// CFC twin of T_SafeOr_Tests: the same tests drawn as CFC diagrams, the way a TwinSAFE project is authored.
    FUNCTION_BLOCK T_SafeOr_Tests_CFC EXTENDS T_SafeCfcTestSuite
    VAR
    // Test_AnyConnectedInputTrueGivesRun
    group_1 : T_SafeGroup;
    fb_1 : T_SafeOr(group := group_1);
    // Test_AllFalseGivesSafe
    group_2 : T_SafeGroup;
    fb_2 : T_SafeOr(group := group_2);
END_VAR

Test_AnyConnectedInputTrueGivesRun();
Test_AllFalseGivesSafe();

METHOD PRIVATE Test_AnyConnectedInputTrueGivesRun
// note: this text did not pass the execution check against the stored diagram
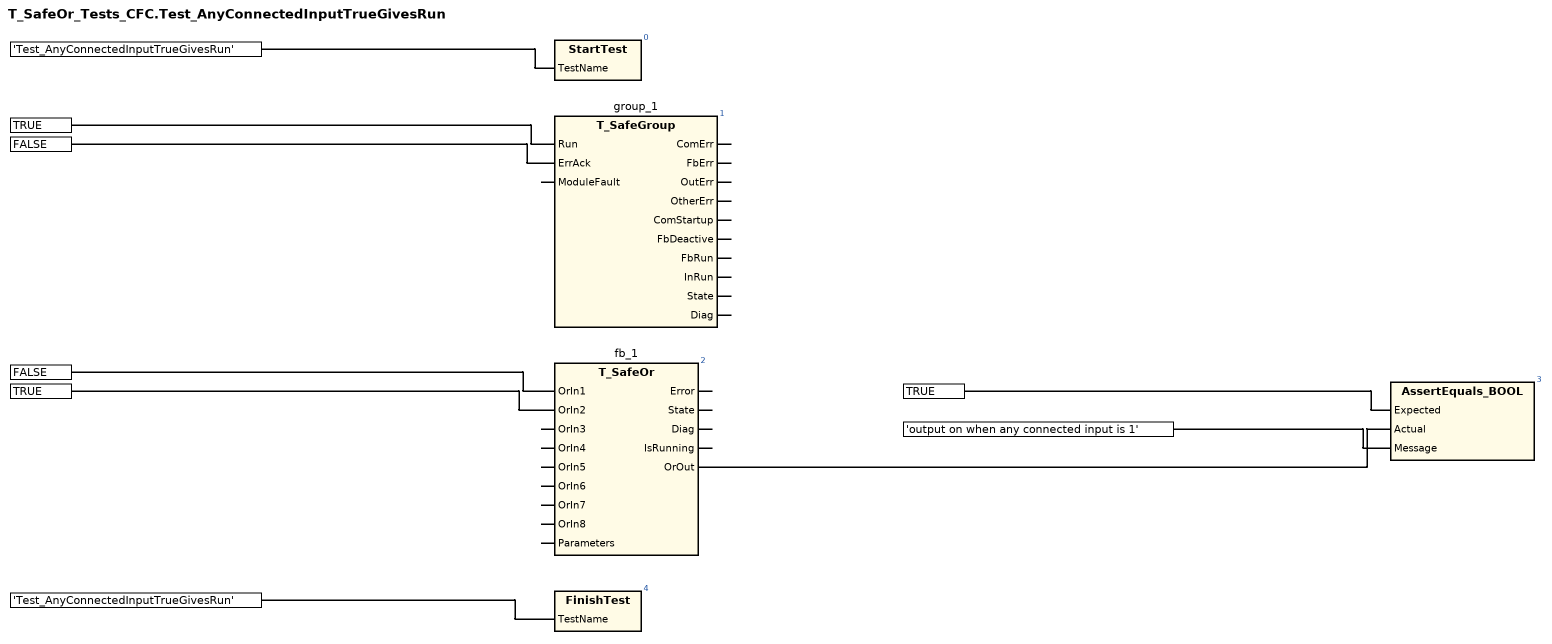
StartTest(TestName := 'Test_AnyConnectedInputTrueGivesRun');
group_1(Run := TRUE, ErrAck := FALSE); // T_SafeGroup
fb_1(OrIn1 := FALSE, OrIn2 := TRUE); // T_SafeOr
AssertEquals_BOOL(Expected := TRUE, Actual := fb_1.OrOut, Message := 'output on when any connected input is 1');
FinishTest(TestName := 'Test_AnyConnectedInputTrueGivesRun');
END_METHOD

METHOD PRIVATE Test_AllFalseGivesSafe
// note: this text did not pass the execution check against the stored diagram
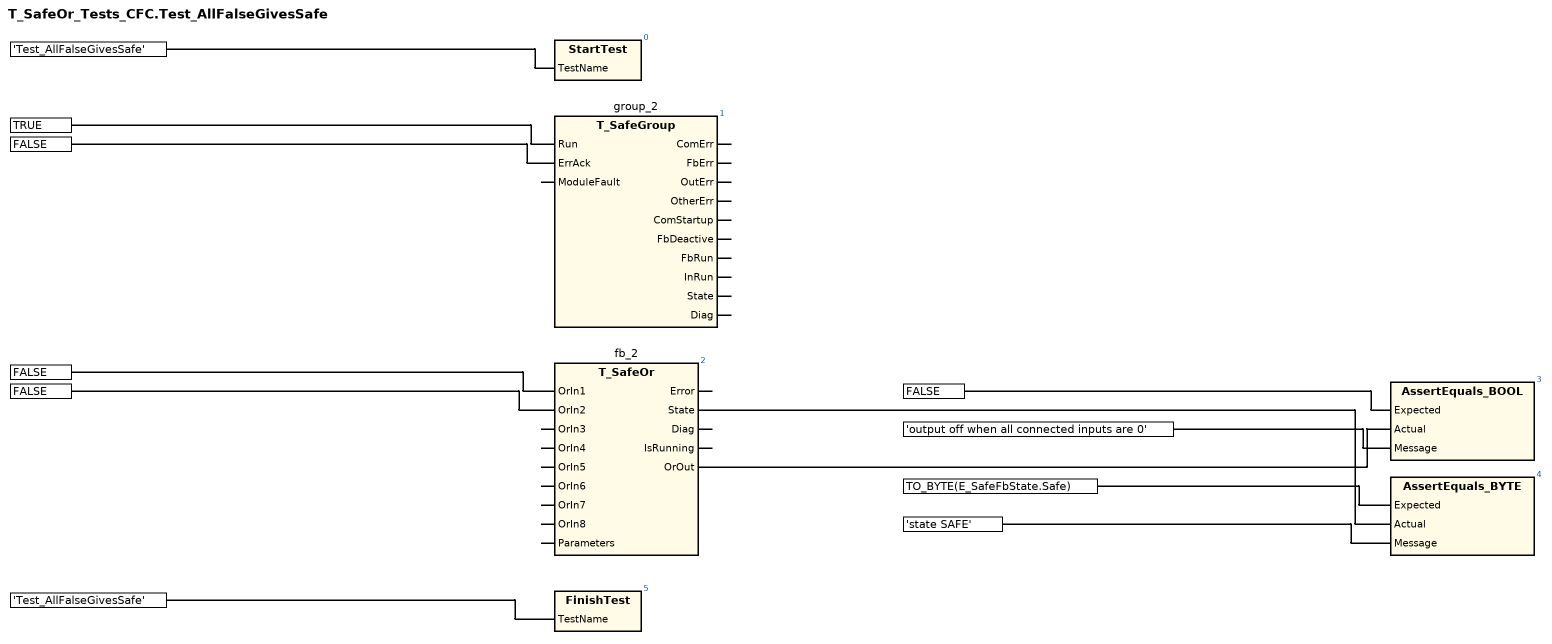
StartTest(TestName := 'Test_AllFalseGivesSafe');
group_2(Run := TRUE, ErrAck := FALSE); // T_SafeGroup
fb_2(OrIn1 := FALSE, OrIn2 := FALSE); // T_SafeOr
AssertEquals_BOOL(Expected := FALSE, Actual := fb_2.OrOut, Message := 'output off when all connected inputs are 0');
AssertEquals_BYTE(Expected := TO_BYTE(E_SafeFbState.Safe), Actual := fb_2.State, Message := 'state SAFE');
FinishTest(TestName := 'Test_AllFalseGivesSafe');
END_METHOD

END_FUNCTION_BLOCK

(* stored: Version 1.1.0.1, ProductVersion 3.1.4026.22
   POU T_SafeOr_Tests_CFC: Id {29568816-f524-5c2f-a8e6-75c0cc1d42f8}, SpecialFunc None
   Method Test_AnyConnectedInputTrueGivesRun: Id {120160bf-b190-5f14-b776-28041d546f05}
   Method Test_AllFalseGivesSafe: Id {a723f035-4c74-58f2-bfac-3e97bae6e99c} *)
